(*
	| return the Process Info from List with {Index} (Base = 0)
*)
METHOD PROTECTED _getProcessInfo : KOSTAL_AF2024_Core_Settings.T_MaxString_UTF8
VAR_INPUT
	IN		: Tc3_IotBase.SJsonValue;
END_VAR

VAR
	_J	: Tc3_IotBase.SJsonValue;
	_uliResult: ULINT;
	_udiResult: UDINT;
	_diResult	: DINT;
	_bResult	: BOOL;
	_sResult	: KOSTAL_AF2024_Core_Settings.T_MaxString_UTF8;
END_VAR

IF IN = 0 												THEN _getProcessInfo:= 'IN Parameter is empty';												RETURN;	END_IF

_ResponseProcess.clear();

_sResp:= _PARSE_JSON(IN, PROCESS_INFO.processInfo, _J);
IF _sResp <> '' THEN	_getProcessInfo:= _sResp;	RETURN; END_IF
IF _J = 0	THEN _getProcessInfo:= '_getProcessInfo - no content availabe';	RETURN;	END_IF

_sResp:= _PARSE_ULINT(_J, PROCESS_INFO.id, _uliResult);
IF _sResp <> '' THEN	_getProcessInfo:= _sResp;	ELSE	_ResponseProcess.id:= _uliResult; END_IF

_sResp:= _PARSE_STRING(_J, PROCESS_INFO.serialNumber, _sResult);
IF _sResp <> '' THEN	_getProcessInfo:= _sResp;	ELSE	_ResponseProcess.serialNumber:= _sResult;	END_IF

_sResp:= _PARSE_STRING(_J, PROCESS_INFO.articleNumber, _sResult);
IF _sResp <> '' THEN	_getProcessInfo:= _sResp;	ELSE	_ResponseProcess.articleNumber:= _sResult;	END_IF

_sResp:= _PARSE_STRING(_J, PROCESS_INFO.timeStamp, _sResult);
IF _sResp <> '' THEN	_getProcessInfo:= _sResp;	ELSE	_ResponseProcess.timeStamp:= _sResult;	END_IF

_sResp:= _PARSE_DINT(_J, PROCESS_INFO.traceId, _diResult);
IF _sResp <> '' THEN	_getProcessInfo:= _sResp;	ELSE	_ResponseProcess.traceId:= _diResult; END_IF

_sResp:= _PARSE_STRING(_J, PROCESS_INFO.process, _sResult);
IF _sResp <> '' THEN	_getProcessInfo:= _sResp;	ELSE	_ResponseProcess.process:= _sResult;	END_IF

_sResp:= _PARSE_BOOL(_J, PROCESS_INFO.result, _bResult);
IF _sResp <> '' THEN	_getProcessInfo:= _sResp;	ELSE	_ResponseProcess.result:= _bResult;	END_IF

_sResp:= _PARSE_STRING(_J, PROCESS_INFO.optionalString_1, _sResult);
IF _sResp <> '' THEN	_getProcessInfo:= _sResp;	ELSE	_ResponseProcess.OptionalStrings_Owner.set(1, _sResult);	END_IF

_sResp:= _PARSE_STRING(_J, PROCESS_INFO.optionalString_2, _sResult);
IF _sResp <> '' THEN	_getProcessInfo:= _sResp;	ELSE	_ResponseProcess.OptionalStrings_Owner.set(2, _sResult);	END_IF

_sResp:= _PARSE_STRING(_J, PROCESS_INFO.optionalString_3, _sResult);
IF _sResp <> '' THEN	_getProcessInfo:= _sResp;	ELSE	_ResponseProcess.OptionalStrings_Owner.set(3, _sResult);	END_IF

_sResp:= _PARSE_STRING(_J, PROCESS_INFO.optionalString_4, _sResult);
IF _sResp <> '' THEN	_getProcessInfo:= _sResp;	ELSE	_ResponseProcess.OptionalStrings_Owner.set(4, _sResult);	END_IF

_sResp:= _PARSE_BOOL(_J, PROCESS_INFO.optionalFlag_1, _bResult);
IF _sResp <> '' THEN	_getProcessInfo:= _sResp;	ELSE	_ResponseProcess.OptionalFlags_Owner.set(1, (_bResult <> 0));	END_IF

_sResp:= _PARSE_BOOL(_J, PROCESS_INFO.optionalFlag_2, _bResult);
IF _sResp <> '' THEN	_getProcessInfo:= _sResp;	ELSE	_ResponseProcess.OptionalFlags_Owner.set(2, (_bResult <> 0));	END_IF

_sResp:= _PARSE_BOOL(_J, PROCESS_INFO.optionalFlag_3, _bResult);
IF _sResp <> '' THEN	_getProcessInfo:= _sResp;	ELSE	_ResponseProcess.OptionalFlags_Owner.set(3, (_bResult <> 0));	END_IF

_sResp:= _PARSE_BOOL(_J, PROCESS_INFO.optionalFlag_4, _bResult);
IF _sResp <> '' THEN	_getProcessInfo:= _sResp;	ELSE	_ResponseProcess.OptionalFlags_Owner.set(4, (_bResult <> 0));	END_IF

_sResp:= _PARSE_BOOL(_J, PROCESS_INFO.optionalFlag_5, _bResult);
IF _sResp <> '' THEN	_getProcessInfo:= _sResp;	ELSE	_ResponseProcess.OptionalFlags_Owner.set(5, (_bResult <> 0));	END_IF

_sResp:= _PARSE_BOOL(_J, PROCESS_INFO.optionalFlag_6, _bResult);
IF _sResp <> '' THEN	_getProcessInfo:= _sResp;	ELSE	_ResponseProcess.OptionalFlags_Owner.set(6, (_bResult <> 0));	END_IF

_sResp:= _PARSE_BOOL(_J, PROCESS_INFO.optionalFlag_7, _bResult);
IF _sResp <> '' THEN	_getProcessInfo:= _sResp;	ELSE	_ResponseProcess.OptionalFlags_Owner.set(7, (_bResult <> 0));	END_IF

_sResp:= _PARSE_BOOL(_J, PROCESS_INFO.optionalFlag_8, _bResult);
IF _sResp <> '' THEN	_getProcessInfo:= _sResp;	ELSE	_ResponseProcess.OptionalFlags_Owner.set(8, (_bResult <> 0));	END_IF
END_METHOD

METHOD PROTECTED _01_Ready : BOOL
VAR_INPUT
END_VAR


IF NOT 	SUPER^._01_Ready() 						THEN	;
ELSIF		_THIS_CALLED = E_PROCESS.idle THEN	_state.clear();	_state.ready:= TRUE;

ELSIF		_THIS_CALLED = E_PROCESS.execute		THEN	

	_THIS_IN_PROCESS:= _THIS_CALLED;	

	_state.clear();	
	_state.busy:= TRUE;

	_selectUrl();

	_step.INC();
	
ELSE

	_state.clear();
	_state.fail:= TRUE;
	_state.description:= Tc2_Standard.WCONCAT("Unknown Process called:", INT_TO_WSTRING(_THIS_CALLED));
	
END_IF
END_METHOD

METHOD PROTECTED _10_getProcessInfo
VAR_INPUT
END_VAR

IF _step.toggle THEN
	;
END_IF

_sResp:= _getProcessInfo(_jsonDoc);

IF _sResp <> '' THEN
	
	_state.clear();
	_state.description:= Tc2_Standard.WCONCAT("Process Info is corrupt;", TO_WSTRING(_sResp));
	_step.set(_ADDRESS_FINISH_FAIL);

ELSE	

	_step.INC();

END_IF
END_METHOD

METHOD PROTECTED _10_processWrite
VAR_INPUT
END_VAR

IF _step.toggle THEN

	_ResponseResult.clear();
	_ResponseProcess.clear();

END_IF

_00_clientCfg();
END_METHOD

METHOD PROTECTED _20_setProcessInfo

VAR
	_JsonArray				: Tc3_IotBase.SJsonValue;
	_JsonArrayMember	: Tc3_IotBase.SJsonValue;

	_s	: KOSTAL_AF2024_Core_Settings.T_MaxString_UTF8;
	_i	: UDINT;
	//_pC	: POINTER TO  KOSTAL_TC3_Components_Linecontrol_I_LC.FB_childSet;
	_di: DINT;
END_VAR

IF _step.toggle THEN
	;
END_IF


_jsonDoc:= _JsonParser.NewDocument();

_s:= _WriteDataDto.serialNumber;
_JsonParser.AddStringMember(_jsondoc, PROCESS_INFO.serialNumber, _s);

_s:= _WriteDataDto.articleNumber;
_JsonParser.AddStringMember(_jsondoc, PROCESS_INFO.articleNumber, _s);

_JsonParser.AddBoolMember(_jsondoc, PROCESS_INFO.result, _WriteDataDto.result);

_JsonParser.AddBoolMember(_jsondoc, PROCESS_INFO.optionalFlag_1, _WriteDataDto.OptionalFlags.get(1));
_JsonParser.AddBoolMember(_jsondoc, PROCESS_INFO.optionalFlag_2, _WriteDataDto.OptionalFlags.get(2));
_JsonParser.AddBoolMember(_jsondoc, PROCESS_INFO.optionalFlag_3, _WriteDataDto.OptionalFlags.get(3));
_JsonParser.AddBoolMember(_jsondoc, PROCESS_INFO.optionalFlag_4, _WriteDataDto.OptionalFlags.get(4));
_JsonParser.AddBoolMember(_jsondoc, PROCESS_INFO.optionalFlag_5, _WriteDataDto.OptionalFlags.get(5));
_JsonParser.AddBoolMember(_jsondoc, PROCESS_INFO.optionalFlag_6, _WriteDataDto.OptionalFlags.get(6));
_JsonParser.AddBoolMember(_jsondoc, PROCESS_INFO.optionalFlag_7, _WriteDataDto.OptionalFlags.get(7));
_JsonParser.AddBoolMember(_jsondoc, PROCESS_INFO.optionalFlag_8, _WriteDataDto.OptionalFlags.get(8));

_s:= _WriteDataDto.OptionalStrings.get(1);
_JsonParser.AddStringMember(_jsondoc, PROCESS_INFO.optionalString_1, _s);

_s:= _WriteDataDto.OptionalStrings.get(2);
_JsonParser.AddStringMember(_jsondoc, PROCESS_INFO.optionalString_2, _s);

_s:= _WriteDataDto.OptionalStrings.get(3);
_JsonParser.AddStringMember(_jsondoc, PROCESS_INFO.optionalString_3, _s);

_s:= _WriteDataDto.OptionalStrings.get(4);
_JsonParser.AddStringMember(_jsondoc, PROCESS_INFO.optionalString_4, _s);

_step.INC();
END_METHOD

(*
|MUST EXTEND
*)
METHOD PROTECTED _selectUrl
END_METHOD

METHOD Execute : BOOL

IF _THIS_CALLED <> E_PROCESS.idle THEN Execute:= FALSE;	RETURN; END_IF

_THIS_CALLED:= E_PROCESS.execute;

_FBmain();

Execute:= _THIS_CALLED = _THIS_IN_PROCESS;
END_METHOD

PROPERTY PUBLIC ResponseProcess : I_T_SingleProcess
GET

ResponseProcess:= _ResponseProcess;
END_GET
END_PROPERTY

PROPERTY ResponseResult : I_T_ResponseResult
GET

ResponseResult := _ResponseResult;
END_GET
END_PROPERTY

PROPERTY PUBLIC WriteDataDto : I_T_WriteCurrentStampDataDto_Owner
GET

WriteDataDto := _WriteDataDto;
END_GET
END_PROPERTY

END_FUNCTION_BLOCK

// 5_POU/WriteProcess/FB_WriteProcess
(*
|MUST EXEND
|
|Extends the base WebService LC with a 
|write
|functionality
*)
FUNCTION_BLOCK PUBLIC FB_WriteProcess EXTENDS _FB_WriteProcess

METHOD PROTECTED _selectUrl


_sUrl:= _UriGet(URL.WRITE_CUR_PROC);

_UrlReplace(_sUrl, URL.PLACEHOLDER_CLIENT_NAME, _ClientName);
_UrlReplace(_sUrl, URL.PLACEHOLDER_CLIENT_PROCESS, _ClientProcess);
END_METHOD

METHOD PROTECTED _FBmain
VAR_INPUT
END_VAR

SUPER^._FBmain();

CASE _step.actual OF

	0:	_01_Ready();
	//
	1:	_10_processWrite();
	2:	_20_setProcessInfo();
	3:	_10_SET(TRUE);
	4:	_10_SET_CTRL();
	5:	_10_GET_ResponseResult(FALSE);
	6:	_10_GET_ResponseResult_CTRL();
	7:	_10_getProcessInfo();
	8:	_10_finishPass();

	100:	_10_finishFail();
ELSE
	
	_99_stepError();
		
END_CASE
END_METHOD

END_FUNCTION_BLOCK

// 5_POU/WriteProcess/FB_WriteProcessWithSM
(*
|MUST EXEND
|
|Extends the base WebService LC with a 
|write
|functionality
*)
FUNCTION_BLOCK PUBLIC FB_WriteProcessWithSM EXTENDS _FB_WriteProcess

VAR

	//======================================================================================
	//Parameter
	//======================================================================================
	
	//_SingleProcess	: FB_SingleProcess;
	_SubModuls			: FB_ListOfSubModule;	

END_VAR

METHOD PROTECTED _20_setSubModules

VAR
	_JsonArrayElement	: Tc3_IotBase.SJsonValue;
	_JsonArray				: Tc3_IotBase.SJsonValue;
	_JsonArrayMember	: Tc3_IotBase.SJsonValue;

	_s	: KOSTAL_AF2024_Core_Settings.T_MaxString_UTF8;
	_udi: UDINT;

END_VAR

IF _step.toggle THEN
	;
END_IF

IF _SubModuls.NumberOfMember = 0 THEN 
	
	_state.clear();
	_state.description:= "No Sub-Modules available";
	_step.set(_ADDRESS_FINISH_FAIL);
	
	RETURN;

END_IF

_JsonArrayElement:= _JsonParser.AddJsonMember(_jsondoc, SUBMODUL_INFO.subModules, '');

IF _JsonArrayElement = 0 THEN 

	_state.clear();
	_state.description:= "Unable to create Sub-Modul Array";
	_step.set(_ADDRESS_FINISH_FAIL);
	
	RETURN;
END_IF

_JsonArray:= _JsonParser.SetArray(_JsonArrayElement, 0);

IF _JsonArray = 0 THEN 

	_state.clear();
	_state.description:= "Unable to create Sub-Modul Array";
	_step.set(_ADDRESS_FINISH_FAIL);
	
	RETURN;
END_IF


FOR _udi:=  1 TO _SubModuls.NumberOfMember DO

	_JsonArrayMember:= 	_JsonParser.PushbackJsonValue(_JsonArray, '');

	//_JsonParser.AddJsonMember(_JsonArray, '', 0);
	
	IF _JsonArrayMember = 0 THEN 
	
		_state.clear();
		_state.description:= "Unable to create Sub-Modul Array";
		_step.set(_ADDRESS_FINISH_FAIL);
		
		RETURN;
	END_IF

	_s:= _SubModuls.Get_I(_udi, 0, 0).articleNumber;
	_JsonParser.AddStringMember(_JsonArrayMember, SUBMODUL_INFO.articleNumber, _s);
	
	_s:= _SubModuls.Get_I(_udi, 0, 0).serialNumber;
	_JsonParser.AddStringMember(_JsonArrayMember, SUBMODUL_INFO.serialNumber, _s);
	
	
END_FOR


_step.INC();
END_METHOD

METHOD PROTECTED _selectUrl


_sUrl:= _UriGet(URL.WRITE_CUR_PROC_WITH_SUBMODULS);

_UrlReplace(_sUrl, URL.PLACEHOLDER_CLIENT_NAME, _ClientName);
_UrlReplace(_sUrl, URL.PLACEHOLDER_CLIENT_PROCESS, _ClientProcess);
END_METHOD

PROPERTY PUBLIC ListOfSubModules : I_ListOfSubModule_Owner
GET

ListOfSubModules := _SubModuls;
END_GET
END_PROPERTY

METHOD PROTECTED _FBmain
VAR_INPUT
END_VAR

SUPER^._FBmain();

CASE _step.actual OF

	0:	_01_Ready();
	//
	1:	_10_processWrite();
	2:	_20_setProcessInfo();
	3:	_20_setSubModules();
	4:	_10_SET(TRUE);
	5:	_10_SET_CTRL();
	6:	_10_GET_ResponseResult(FALSE);
	7:	_10_GET_ResponseResult_CTRL();
	8:	_10_getProcessInfo();
	9:	_10_finishPass();

	100:	_10_finishFail();
ELSE
	
	_99_stepError();
		
END_CASE
END_METHOD

END_FUNCTION_BLOCK

// Project Information/F_GetCompany
// This function has been automatically generated from the project information.
{attribute 'signature_flag' := '1073741824'}
{attribute 'TcGenerated'}
{attribute 'no-analysis'}
FUNCTION F_GetCompany : WSTRING
VAR_INPUT
	
END_VAR

F_GetCompany := "KOSTAL GmbH & Co.KG";

END_FUNCTION
